FUNCTION_BLOCK UCT_Equipamento_HMI (* Service Interface Function Block Type *)
  (* Standard: 61499-2 *)
  (* Version 1.5, 03/11/2026, Hidryco, Hidryco, 1.5: nomes no padrao do Citect (CMD_MANUAL, STP_VELOCIDADE, CMD_INTERMITENTE, HABILITA_REVERSAO, STS_HORIMETRO_HOR). IHM de um equipamento da UCT (nomes dos CATs Peneira_Rotativa/Bomba_Higienizacao/Rosca...) *)
  PACKAGE Hidryco.HidrycoLib;
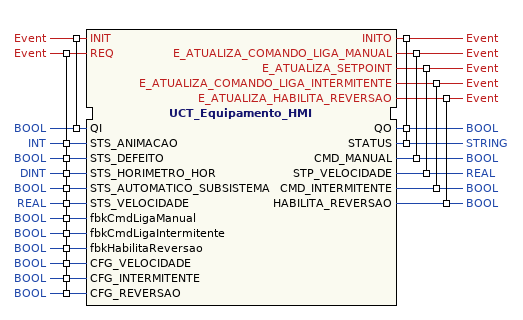
  EVENT_INPUT
    INIT WITH QI;
    REQ WITH STS_ANIMACAO, STS_DEFEITO, STS_HORIMETRO_HOR, STS_AUTOMATICO_SUBSISTEMA, STS_VELOCIDADE, fbkCmdLigaManual, fbkCmdLigaIntermitente, fbkHabilitaReversao, CFG_VELOCIDADE, CFG_INTERMITENTE, CFG_REVERSAO; (* Atualizacao de status *)
  END_EVENT
  EVENT_OUTPUT
    INITO WITH QO, STATUS;
    E_ATUALIZA_COMANDO_LIGA_MANUAL WITH CMD_MANUAL;
    E_ATUALIZA_SETPOINT WITH STP_VELOCIDADE;
    E_ATUALIZA_COMANDO_LIGA_INTERMITENTE WITH CMD_INTERMITENTE;
    E_ATUALIZA_HABILITA_REVERSAO WITH HABILITA_REVERSAO;
  END_EVENT
  VAR_INPUT
    QI : BOOL;
    STS_ANIMACAO : INT; (* Estado do equipamento na UCT: 0 desligado, 1 ligado, 2 falha, 3 manutencao, 4 sem comunicacao *)
    STS_DEFEITO : BOOL; (* Defeito do equipamento (palavra 40081 da UCT) *)
    STS_HORIMETRO_HOR : DINT; (* Horimetro do equipamento (h, lido da UCT) *)
    STS_AUTOMATICO_SUBSISTEMA : BOOL; (* Subsistema do equipamento em automatico (comandos manuais bloqueados) *)
    STS_VELOCIDADE : REAL; (* Velocidade ajustada na UCT (Hz) *)
    fbkCmdLigaManual : BOOL; (* Comando liga em vigor na UCT *)
    fbkCmdLigaIntermitente : BOOL; (* Modo intermitente em vigor na UCT *)
    fbkHabilitaReversao : BOOL; (* Reversao habilitada na UCT *)
    CFG_VELOCIDADE : BOOL; (* TRUE = equipamento com ajuste de velocidade *)
    CFG_INTERMITENTE : BOOL; (* TRUE = equipamento com modo intermitente *)
    CFG_REVERSAO : BOOL; (* TRUE = equipamento com reversao *)
  END_VAR
  VAR_OUTPUT
    QO : BOOL; (* Event Output Qualifier *)
    STATUS : STRING; (* Service Status *)
    CMD_MANUAL : BOOL; (* IHM: liga (TRUE) / desliga (FALSE) em manual *)
    STP_VELOCIDADE : REAL; (* IHM: velocidade (Hz) *)
    CMD_INTERMITENTE : BOOL; (* IHM: liga (TRUE) / desliga (FALSE) o intermitente *)
    HABILITA_REVERSAO : BOOL; (* IHM: habilita (TRUE) / desabilita (FALSE) a reversao *)
  END_VAR
  SERVICE /
    SEQUENCE 
    END_SEQUENCE
  END_SERVICE
END_FUNCTION_BLOCK
